// LS Electric XG5000 project: REMRES
// PLC LSPLC

PROGRAM NewProgram (task: 스캔 프로그램)

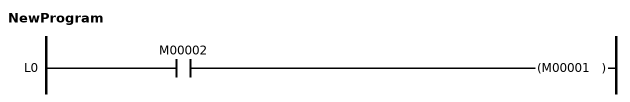
; L0
LOAD      M00002
OUT       M00001